(* CODESYS project i_linearaxis.library
   DefaultNamespace: KOSTAL.TC3.Device.Axis.I_LinearAxis
   DocFormat: reStructuredText
   Description: Application interface for linear axis control:
      - Common base interface
      - Jog mode interface for 1D, 2D and 3D axis
      - Position control interface for 1D, 2D and 3D axis
      - Record mode interface (1D, 2D and 3D mode to be handled in the driver)
   Author: Martin Hundt
   Title: KOSTAL.TC3.Device.Axis.I_LinearAxis
   Version: 2019.1.0.0
   Company: KOSTAL GmbH & Co.KG
   Placeholder: KOSTAL.TC3.Device.Axis.I_LinearAxis

Project tree, tasks and I/O mapping:
  libraries: KOSTAL.TC3.Core.plcResponse, * (KOSTAL GmbH & Co.KG)
  Interface/
    1D/
      interface I_LinearAxis_jog: IlinearAxis_JogNegative_X, IlinearAxis_JogPositive_X
      interface I_LinearAxis_position: IlinearAxis_MoveToPosition, IlinearAxis_PositionAct
    2D/
      interface I_LinearAxis_jog_2D: IlinearAxis_JogNegative_Y, IlinearAxis_JogPositive_Y
      interface I_LinearAxis_position2D: IlinearAxis_MoveToPosition, IlinearAxis_PositionAct_X, IlinearAxis_PositionAct_Y
    3D/
      interface I_LinearAxis_jog_3D: IlinearAxis_JogNegative_Z, IlinearAxis_JogPositive_Z
      interface I_LinearAxis_position3D: IlinearAxis_MoveToPosition, IlinearAxis_PositionAct_X, IlinearAxis_PositionAct_Y, IlinearAxis_PositionAct_Z
    interface I_LinearAxis_base: IlinearAxis_acceleration, IlinearAxis_deceleration, IlinearAxis_Fault, IlinearAxis_Homing, IlinearAxis_Off, IlinearAxis_On, IlinearAxis_Release, IlinearAxis_ResetFault, IlinearAxis_Speed, IlinearAxis_State
    interface I_LinearAxis_record: IlinearAxis_MoveRecord
  Project Information/
    function F_GetCompany [ST]
    function F_GetTitle [ST]
    function F_GetVersion [ST]
  Version/
    global variables Global_Version
*)

// Version/Global_Version
{attribute 'TcGenerated'}
{attribute 'no-analysis'}
{attribute 'linkalways'}
// This function has been automatically generated from the project information.
VAR_GLOBAL CONSTANT
	{attribute 'const_non_replaced'}
	stLibVersion_KOSTAL_TC3_Device_Axis_I_LinearAxis : ST_LibVersion := (iMajor := 2019, iMinor := 1, iBuild := 0, iRevision := 0, nFlags := 0, sVersion := '2019.1.0.0');
END_VAR

// Interface/1D/I_LinearAxis_jog
(*
:Author: Martin Hundt <m.hundt@kostal.com>, 
:Date: 2020-11-30

Function
========
| Control linear axis in jog mode

Methods
=======
| JogNegative_X/JogPositive_X: Move axis in positive or nagative direction. Speed and acceleration to be defined via properties in the base class.

*)
INTERFACE I_LinearAxis_jog EXTENDS I_LinearAxis_base

METHOD IlinearAxis_JogNegative_X
VAR_INPUT
END_VAR
END_METHOD

METHOD IlinearAxis_JogPositive_X
VAR_INPUT
END_VAR
END_METHOD

END_INTERFACE

// Interface/I_LinearAxis_base
(*
:Author: Martin Hundt <m.hundt@kostal.com>, 
:Date: 2020-11-30

Function
========
| Base class to control linear axis
| To be extended with jog, position or record interface


Properties
==========
| acceleration / IlinearAxis_deceleration: Acceleration and deceleration in mm/s²
| Speed: Axis velocity in mm/s
| State: Feedback of device's state (see main documentation)
| Fault: TRUE in case of device fault. Error message to be found in state.description

Methods
=======
| Notes: 
| - If a certain device does not support a function (e.g. homing, the implemented method shall just feed back sucess
| - Some methods have a boolean return value. Set it TRUE if the method succeeded, but also use the finish and pass/fail bits of the state property!
| On/Off: Switch axis power on or off
| Release: release axis movement (e.g. release brakes)
| Homing: Carry out the axis homing sequence (device dependent)
| ResetFault

Usage sample:
=============
See actual device drivers that implement the interface
*)
INTERFACE I_LinearAxis_base

PROPERTY IlinearAxis_acceleration : REAL
GET
END_GET
SET
END_SET
END_PROPERTY

PROPERTY IlinearAxis_deceleration : REAL
GET
END_GET
SET
END_SET
END_PROPERTY

PROPERTY IlinearAxis_Fault : BOOL
GET
END_GET
END_PROPERTY

METHOD IlinearAxis_Homing : BOOL
VAR_INPUT
END_VAR
END_METHOD

METHOD IlinearAxis_Off : BOOL
END_METHOD

METHOD IlinearAxis_On : BOOL
END_METHOD

METHOD IlinearAxis_Release : BOOL
VAR_INPUT
	release : BOOL;
END_VAR
END_METHOD

METHOD IlinearAxis_ResetFault  : BOOL
END_METHOD

PROPERTY IlinearAxis_Speed : REAL
GET
END_GET
SET
END_SET
END_PROPERTY

PROPERTY IlinearAxis_State : REFERENCE TO KOSTAL_TC3_Core_plcResponse.FB_PlcResponse;
GET
END_GET
END_PROPERTY

END_INTERFACE

// Interface/1D/I_LinearAxis_position
(*
:Author: Martin Hundt <m.hundt@kostal.com>, 
:Date: 2020-11-30

Function
========
| Control linear axis in positioning mode

Methods
=======
| MoveToPosition(REAL position): Move axis to given position, Unit: mm. Speed and acceleration to be defined via properties in the base class.

Properties
==========
| PositionAct: Actual position of the axis in mm
*)

INTERFACE I_LinearAxis_position EXTENDS I_LinearAxis_base


//Move to given position
METHOD IlinearAxis_MoveToPosition
VAR_INPUT
	position	: REAL;
END_VAR
END_METHOD

PROPERTY IlinearAxis_PositionAct : Real
GET
END_GET
END_PROPERTY

END_INTERFACE

// Interface/2D/I_LinearAxis_jog_2D
(*
:Author: Martin Hundt <m.hundt@kostal.com>, 
:Date: 2020-11-30

Function
========
| Extension of IlinearAxis_jog to control 2D axis

*)
INTERFACE I_LinearAxis_jog_2D EXTENDS I_LinearAxis_jog

METHOD IlinearAxis_JogNegative_Y
VAR_INPUT
END_VAR
END_METHOD

METHOD IlinearAxis_JogPositive_Y
VAR_INPUT
END_VAR
END_METHOD

END_INTERFACE

// Interface/2D/I_LinearAxis_position2D
(*
:Author: Martin Hundt <m.hundt@kostal.com>, 
:Date: 2020-11-30

Function
========
| Extension of IlinearAxis_position to control 2D axis

*)
INTERFACE I_LinearAxis_position2D EXTENDS I_LinearAxis_base


//Move to given position
METHOD IlinearAxis_MoveToPosition
VAR_INPUT
	positionX	: REAL;
	positionY	: REAL;
END_VAR
END_METHOD

PROPERTY IlinearAxis_PositionAct_X : Real
GET
END_GET
END_PROPERTY

PROPERTY IlinearAxis_PositionAct_Y : Real
GET
END_GET
END_PROPERTY

END_INTERFACE

// Interface/3D/I_LinearAxis_jog_3D
(*
:Author: Martin Hundt <m.hundt@kostal.com>, 
:Date: 2020-11-30

Function
========
| Extension of IlinearAxis_jog to control 3D axis

*)
INTERFACE I_LinearAxis_jog_3D EXTENDS I_LinearAxis_jog_2D

METHOD IlinearAxis_JogNegative_Z
VAR_INPUT
END_VAR
END_METHOD

METHOD IlinearAxis_JogPositive_Z
VAR_INPUT
END_VAR
END_METHOD

END_INTERFACE

// Interface/3D/I_LinearAxis_position3D
(*
:Author: Martin Hundt <m.hundt@kostal.com>, 
:Date: 2020-11-30

Function
========
| Extension of IlinearAxis_position to control 3D axis

*)
INTERFACE I_LinearAxis_position3D EXTENDS I_LinearAxis_base


//Move to given position
METHOD IlinearAxis_MoveToPosition
VAR_INPUT
	positionX	: REAL;
	positionY	: REAL;
	positionZ	: REAL;
END_VAR
END_METHOD

PROPERTY IlinearAxis_PositionAct_X : Real
GET
END_GET
END_PROPERTY

PROPERTY IlinearAxis_PositionAct_Y : Real
GET
END_GET
END_PROPERTY

PROPERTY IlinearAxis_PositionAct_Z : Real
GET
END_GET
END_PROPERTY

END_INTERFACE

// Interface/I_LinearAxis_record
(*
:Author: Martin Hundt <m.hundt@kostal.com>, 
:Date: 2020-11-30

Function
========
| Control linear axis in record mode (positions and other movement parameters are stored in the axis device)
| In case the parameter set also contains values from the interface base, the interface values shall be ignored

Methods
=======
| MoveRecord (UINT recordNo): Carry out movement of given parameter set

*)

INTERFACE I_LinearAxis_record EXTENDS I_LinearAxis_base

METHOD IlinearAxis_MoveRecord 
VAR_INPUT
	recordNo	: UINT;
END_VAR
END_METHOD

END_INTERFACE

// Project Information/F_GetCompany
// This function has been automatically generated from the project information.
{attribute 'signature_flag' := '1073741824'}
{attribute 'TcGenerated'}
{attribute 'no-analysis'}
FUNCTION F_GetCompany : WSTRING
VAR_INPUT
	
END_VAR

F_GetCompany := "KOSTAL GmbH & Co.KG";

END_FUNCTION

// Project Information/F_GetTitle
// This function has been automatically generated from the project information.
{attribute 'signature_flag' := '1073741824'}
{attribute 'TcGenerated'}
{attribute 'no-analysis'}
FUNCTION F_GetTitle : WSTRING
VAR_INPUT
	
END_VAR

F_GetTitle := "KOSTAL.TC3.Device.Axis.I_LinearAxis";

END_FUNCTION

// Project Information/F_GetVersion
// This function has been automatically generated from the project information.
{attribute 'signature_flag' := '1073741824'}
{attribute 'TcGenerated'}
{attribute 'no-analysis'}
FUNCTION F_GetVersion : ST_LibVersion
VAR_INPUT
	
END_VAR

F_GetVersion.iMajor := 2019;
F_GetVersion.iMinor := 1;
F_GetVersion.iBuild := 0;
F_GetVersion.iRevision := 0;

END_FUNCTION
